(* IEC 61131-3 sources: weg-plc500-nodered-ml-pipeline/plc/src, 5 files *)

(* ---- GVL_Modbus.st ---- *)
{attribute 'qualified_only'}
VAR_GLOBAL
  (* ===================================================================== *)
  (* 1. E/S Fisicas Nativas - WEG PLC500 Local_IO (24 Vcc PNP)             *)
  (* ===================================================================== *)
  xRaw_DI0_Presenca   AT %IX0.0 : BOOL;          (* B1_SensPresenca - Contato NA *)
  xRaw_DI1_NivelAlto  AT %IX0.1 : BOOL;          (* B2_SensNivelAlto - Contato NA *)
  xRaw_DI2_Sobretemp  AT %IX0.2 : BOOL;          (* B3_SensSobretemp - Contato NA *)
  xRaw_DI3_Emergencia AT %IX0.3 : BOOL;          (* B4_Emergencia - Contato NF fail-safe (FALSE = emerg./fio partido) *)

  xDO0_Motor          AT %QX0.0 : BOOL := FALSE; (* L1_AtuMotor - LED Verde *)
  xDO1_Valvula        AT %QX0.1 : BOOL := FALSE; (* L2_AtuValvula - LED Amarelo *)
  xDO2_Alarme         AT %QX0.2 : BOOL := FALSE; (* L3_SinalAlarme - LED Vermelho *)
  xDO3_StatusOper     AT %QX0.3 : BOOL := FALSE; (* L4_StatusOper - LED Branco *)

  (* ===================================================================== *)
  (* 2. Discrete Inputs - Modbus FC02 (Enderecos base zero 0..5)           *)
  (* ===================================================================== *)
  xDI_Presenca : BOOL := FALSE; (* DI[0]: Estado filtrado (TON 50 ms) de B1_SensPresenca *)
  xDI_NivelAlto : BOOL := FALSE; (* DI[1]: Estado filtrado (TON 50 ms) de B2_SensNivelAlto *)
  xDI_Sobretemp : BOOL := FALSE; (* DI[2]: Estado filtrado (TON 50 ms) de B3_SensSobretemp *)
  xDI_EmergenciaOK : BOOL := TRUE; (* DI[3]: Estado imediato NF de B4_Emergencia (TRUE em repouso; FALSE = emergencia) *)
  xFlag_EmergTravada : BOOL := FALSE; (* DI[4]: 1 = emergencia travada aguardando rearme seguro *)
  xFlag_WatchdogAtivo : BOOL := FALSE; (* DI[5]: 1 = heartbeat estagnado > uiTimeout_WD_ms *)

  (* ===================================================================== *)
  (* 3. Coils - Modbus FC01/05/15 (Enderecos base zero 0..4)               *)
  (* ===================================================================== *)
  xCmd_Motor : BOOL := FALSE; (* Coil[0]: Comando remoto para L1_AtuMotor (DO0) *)
  xCmd_Valvula : BOOL := FALSE; (* Coil[1]: Comando remoto para L2_AtuValvula (DO1) *)
  xCmd_Alarme : BOOL := FALSE; (* Coil[2]: Comando remoto para L3_SinalAlarme (DO2) *)
  xCmd_ResetFalha : BOOL := FALSE; (* Coil[3]: Pulso de rearme (borda de subida; valido se DI3=1 e DI2=0) *)
  xCmd_HabRemoto : BOOL := FALSE; (* Coil[4]: 1 = habilita modo automatico supervisionado *)

  (* ===================================================================== *)
  (* 4. Input Registers - Modbus FC04 (Enderecos base zero 0..7)           *)
  (* ===================================================================== *)
  uiCnt_Presenca : UINT := 0; (* IR[0]: Contador modular 16 bits de B1 (0..65535) *)
  uiCnt_NivelAlto : UINT := 0; (* IR[1]: Contador modular 16 bits de B2 (0..65535) *)
  uiCnt_Sobretemp : UINT := 0; (* IR[2]: Contador modular 16 bits de B3 (0..65535) *)
  uiCnt_Emergencia : UINT := 0; (* IR[3]: Contador modular 16 bits de eventos em B4 (0..65535) *)
  uiEstado_CLP : UINT := 0; (* IR[4]: 0=INIT, 1=NORMAL_AUTO, 2=ALERTA, 3=MODO_DEGRADADO, 4=EMERGENCIA_TRAV *)
  wMascara_DO_Real : WORD := 0; (* IR[5]: Bitmask das saidas fisicas (bit0=DO0..bit3=DO3) *)
  uiEcho_Heartbeat : UINT := 0; (* IR[6]: Eco do ultimo valor de heartbeat recebido *)
  uiCod_Intertrav : UINT := 0; (* IR[7]: 0=Nenhum, 1=Emergencia, 2=Sobretemp, 3=Watchdog *)

  (* ===================================================================== *)
  (* 5. Holding Registers - Modbus FC03/06/16 (Enderecos base zero 0..3)   *)
  (* ===================================================================== *)
  uiHeartbeat_Sup : UINT := 0; (* HR[0]: Heartbeat ciclico 1..65535 (aliases de compatibilidade: uiHeartbeat_NR, uiHeartbeat_N8N) *)
  uiTimeout_WD_ms : UINT := 5000; (* HR[1]: Timeout do watchdog em ms [2000..30000], padrao 5000 *)
  uiSeveridade_IA : UINT := 0; (* HR[2]: 0=NORMAL, 1=ATENCAO, 2=CRITICO, 3=EMERGENCIA *)
  uiVersao_Mapa : UINT := 100; (* HR[3]: Versao fixa do contrato Modbus (100 = v1.0) *)
END_VAR

(* ---- FB_DebounceCounter.st ---- *)
FUNCTION_BLOCK FB_DebounceCounter
VAR_INPUT
  xRawInput       : BOOL;           (* Sinal fisico bruto (%IX0.x) *)
  xEnableDebounce : BOOL := TRUE;   (* TRUE = filtro TON (DI0..DI2); FALSE = imediato sem retardo (DI3 NF) *)
  tDebounceTime   : TIME := T#50MS; (* Tempo de estabilizacao de contato *)
  xCountOnFalling : BOOL := FALSE;  (* FALSE = borda de subida (NA); TRUE = borda de descida / NOT (NF DI3) *)
END_VAR
VAR_OUTPUT
  xFiltered       : BOOL := FALSE;  (* Estado filtrado (ou direto para DI3) *)
END_VAR
VAR_IN_OUT
  uiCounter       : UINT;           (* Contador modular 16 bits (wrap natural 65535 -> 0) *)
END_VAR
VAR
  tonDebounce     : STANDARD.TON;
  rtEdge          : STANDARD.R_TRIG;
  xEdgeSignal     : BOOL := FALSE;
END_VAR

IF xEnableDebounce THEN
  tonDebounce(IN := xRawInput, PT := tDebounceTime);
  xFiltered := tonDebounce.Q;
ELSE
  (* Entrada fail-safe DI3 atua sem retardo no primeiro ciclo de varredura *)
  xFiltered := xRawInput;
END_IF;

IF xCountOnFalling THEN
  xEdgeSignal := NOT xFiltered;
ELSE
  xEdgeSignal := xFiltered;
END_IF;

rtEdge(CLK := xEdgeSignal);
IF rtEdge.Q THEN
  uiCounter := uiCounter + 1;
END_IF;
END_FUNCTION_BLOCK

(* ---- FB_SafetyInterlock.st ---- *)
FUNCTION_BLOCK FB_SafetyInterlock
VAR_INPUT
  xDI_EmergenciaOK    : BOOL; (* DI[3]: Contato NF; FALSE = emergencia ativa / fio partido *)
  xDI_Sobretemp       : BOOL; (* DI[2]: Termostato filtrado *)
  xDI_NivelAlto       : BOOL; (* DI[1]: Nivel alto filtrado *)
  xFlag_WatchdogAtivo : BOOL; (* DI[5]: Watchdog expirado *)
  xCmd_Motor          : BOOL; (* Coil[0] *)
  xCmd_Valvula        : BOOL; (* Coil[1] *)
  xCmd_Alarme         : BOOL; (* Coil[2] *)
  xCmd_ResetFalha     : BOOL; (* Coil[3] *)
  xCmd_HabRemoto      : BOOL; (* Coil[4] *)
  uiSeveridade_IA     : UINT; (* HR[2] *)
END_VAR
VAR_OUTPUT
  xFlag_EmergTravada  : BOOL := FALSE; (* DI[4] *)
  uiEstado_CLP        : UINT := 0;     (* IR[4] *)
  uiCod_Intertrav     : UINT := 0;     (* IR[7] *)
  xDO0_Motor          : BOOL := FALSE; (* %QX0.0 *)
  xDO1_Valvula        : BOOL := FALSE; (* %QX0.1 *)
  xDO2_Alarme         : BOOL := FALSE; (* %QX0.2 *)
  xDO3_StatusOper     : BOOL := FALSE; (* %QX0.3 *)
  wMascara_DO_Real    : WORD := 0;     (* IR[5] *)
END_VAR
VAR
  rtResetFalha        : STANDARD.R_TRIG;
END_VAR

(* Deteccao de borda de subida no comando de rearme executada em todo ciclo sem mutar Coil[3] *)
rtResetFalha(CLK := xCmd_ResetFalha);

(* Travamento de emergencia fail-safe e rearme seguro *)
IF NOT xDI_EmergenciaOK THEN
  xFlag_EmergTravada := TRUE;
ELSIF xCmd_ResetFalha AND rtResetFalha.Q AND xDI_EmergenciaOK AND NOT xDI_Sobretemp THEN
  xFlag_EmergTravada := FALSE;
END_IF;

(* Maquina de estados e intertravamento local com precedencia estrita *)
IF xFlag_EmergTravada THEN
  uiEstado_CLP    := 4;
  uiCod_Intertrav := 1;
  xDO0_Motor      := FALSE;
  xDO1_Valvula    := FALSE;
  xDO2_Alarme     := TRUE;
  xDO3_StatusOper := FALSE;
ELSIF xDI_Sobretemp THEN
  uiEstado_CLP    := 2;
  uiCod_Intertrav := 2;
  xDO0_Motor      := FALSE;
  xDO1_Valvula    := TRUE;
  xDO2_Alarme     := TRUE;
  (* Reconciliacao 04_implementacao_clp.tex:141 vs :165/PROJECT.md:110: exige modo remoto ativo alem de watchdog saudavel *)
  xDO3_StatusOper := (NOT xFlag_WatchdogAtivo) AND xCmd_HabRemoto;
ELSIF xFlag_WatchdogAtivo THEN
  uiEstado_CLP    := 3;
  uiCod_Intertrav := 3;
  xDO0_Motor      := FALSE;
  xDO1_Valvula    := xDI_NivelAlto;
  xDO2_Alarme     := TRUE;
  xDO3_StatusOper := FALSE;
ELSIF xCmd_HabRemoto THEN
  uiCod_Intertrav := 0;
  uiEstado_CLP    := SEL((uiSeveridade_IA > 0) OR xDI_NivelAlto, UINT#1, UINT#2);
  xDO0_Motor      := xCmd_Motor;
  xDO1_Valvula    := xCmd_Valvula OR xDI_NivelAlto;
  xDO2_Alarme     := xCmd_Alarme OR (uiSeveridade_IA >= 2);
  xDO3_StatusOper := TRUE;
ELSE
  uiEstado_CLP    := 0;
  uiCod_Intertrav := 0;
  xDO0_Motor      := FALSE;
  xDO1_Valvula    := FALSE;
  xDO2_Alarme     := FALSE;
  xDO3_StatusOper := FALSE;
END_IF;

(* Espelhamento das saidas fisicas reais em bitmask (IR[5]) *)
wMascara_DO_Real := BOOL_TO_WORD(xDO0_Motor)
                 OR SHL(BOOL_TO_WORD(xDO1_Valvula), 1)
                 OR SHL(BOOL_TO_WORD(xDO2_Alarme), 2)
                 OR SHL(BOOL_TO_WORD(xDO3_StatusOper), 3);
END_FUNCTION_BLOCK

(* ---- FB_WatchdogHeartbeat.st ---- *)
FUNCTION_BLOCK FB_WatchdogHeartbeat
VAR_INPUT
  uiHeartbeat     : UINT;          (* HR[0]: uiHeartbeat_Sup (aliases: uiHeartbeat_NR, uiHeartbeat_N8N) *)
  uiTimeoutMs     : UINT;          (* HR[1]: uiTimeout_WD_ms [2000..30000] *)
END_VAR
VAR_OUTPUT
  uiEcho_Heartbeat    : UINT := 0;     (* IR[6]: uiEcho_Heartbeat *)
  xFlag_WatchdogAtivo : BOOL := FALSE; (* DI[5]: xFlag_WatchdogAtivo *)
  tActiveLimit        : TIME := T#5S;  (* Limiar efetivo em TIME *)
END_VAR
VAR
  tonWatchdog     : STANDARD.TON;
  uiLastHeartbeat : UINT := 0;
END_VAR

IF (uiTimeoutMs >= 2000) AND (uiTimeoutMs <= 30000) THEN
  tActiveLimit := UINT_TO_TIME(uiTimeoutMs);
ELSE
  tActiveLimit := T#5S;
END_IF;

(* Avaliar TON ANTES de atualizar uiLastHeartbeat para reiniciar por 1 ciclo na mudanca *)
tonWatchdog(
  IN := (uiHeartbeat = uiLastHeartbeat),
  PT := tActiveLimit
);

IF uiHeartbeat <> uiLastHeartbeat THEN
  uiLastHeartbeat := uiHeartbeat;
  uiEcho_Heartbeat := uiHeartbeat;
END_IF;

xFlag_WatchdogAtivo := tonWatchdog.Q;
END_FUNCTION_BLOCK

(* ---- PLC_PRG.st ---- *)
PROGRAM PLC_PRG
VAR
  fbDebPresenca : FB_DebounceCounter;
  fbDebNivel    : FB_DebounceCounter;
  fbDebTemp     : FB_DebounceCounter;
  rtEmergencia  : STANDARD.R_TRIG;
  fbWatchdog    : FB_WatchdogHeartbeat;
  fbInterlock   : FB_SafetyInterlock;
END_VAR

(* 1 & 2. Debounce (50 ms em DI0..DI2, imediato NF em DI3) e contadores modulares 16 bits *)
GVL_Modbus.xRaw_DI0_Presenca := %IX0.0;
fbDebPresenca(
  xRawInput       := %IX0.0,
  xEnableDebounce := TRUE,
  tDebounceTime   := T#50MS,
  xCountOnFalling := FALSE,
  uiCounter       := GVL_Modbus.uiCnt_Presenca
);
GVL_Modbus.xDI_Presenca := fbDebPresenca.xFiltered;

GVL_Modbus.xRaw_DI1_NivelAlto := %IX0.1;
fbDebNivel(
  xRawInput       := %IX0.1,
  xEnableDebounce := TRUE,
  tDebounceTime   := T#50MS,
  xCountOnFalling := FALSE,
  uiCounter       := GVL_Modbus.uiCnt_NivelAlto
);
GVL_Modbus.xDI_NivelAlto := fbDebNivel.xFiltered;

GVL_Modbus.xRaw_DI2_Sobretemp := %IX0.2;
fbDebTemp(
  xRawInput       := %IX0.2,
  xEnableDebounce := TRUE,
  tDebounceTime   := T#50MS,
  xCountOnFalling := FALSE,
  uiCounter       := GVL_Modbus.uiCnt_Sobretemp
);
GVL_Modbus.xDI_Sobretemp := fbDebTemp.xFiltered;

GVL_Modbus.xRaw_DI3_Emergencia := %IX0.3;
GVL_Modbus.xDI_EmergenciaOK := %IX0.3;
rtEmergencia(CLK := NOT GVL_Modbus.xDI_EmergenciaOK);
IF rtEmergencia.Q THEN
  GVL_Modbus.uiCnt_Emergencia := GVL_Modbus.uiCnt_Emergencia + 1;
END_IF;

(* 3. Supervisao de enlace Modbus TCP/IP (Watchdog via HR[0]/HR[1]) *)
fbWatchdog(
  uiHeartbeat         := GVL_Modbus.uiHeartbeat_Sup,
  uiTimeoutMs         := GVL_Modbus.uiTimeout_WD_ms,
  uiEcho_Heartbeat    => GVL_Modbus.uiEcho_Heartbeat,
  xFlag_WatchdogAtivo => GVL_Modbus.xFlag_WatchdogAtivo
);

(* 4, 5 & 6a. Travamento fail-safe, FSM com precedencia estrita e wMascara_DO_Real *)
fbInterlock(
  xDI_EmergenciaOK    := GVL_Modbus.xDI_EmergenciaOK,
  xDI_Sobretemp       := GVL_Modbus.xDI_Sobretemp,
  xDI_NivelAlto       := GVL_Modbus.xDI_NivelAlto,
  xFlag_WatchdogAtivo := GVL_Modbus.xFlag_WatchdogAtivo,
  xCmd_Motor          := GVL_Modbus.xCmd_Motor,
  xCmd_Valvula        := GVL_Modbus.xCmd_Valvula,
  xCmd_Alarme         := GVL_Modbus.xCmd_Alarme,
  xCmd_ResetFalha     := GVL_Modbus.xCmd_ResetFalha,
  xCmd_HabRemoto      := GVL_Modbus.xCmd_HabRemoto,
  uiSeveridade_IA     := GVL_Modbus.uiSeveridade_IA,
  xFlag_EmergTravada  => GVL_Modbus.xFlag_EmergTravada,
  uiEstado_CLP        => GVL_Modbus.uiEstado_CLP,
  uiCod_Intertrav     => GVL_Modbus.uiCod_Intertrav,
  xDO0_Motor          => GVL_Modbus.xDO0_Motor,
  xDO1_Valvula        => GVL_Modbus.xDO1_Valvula,
  xDO2_Alarme         => GVL_Modbus.xDO2_Alarme,
  xDO3_StatusOper     => GVL_Modbus.xDO3_StatusOper,
  wMascara_DO_Real    => GVL_Modbus.wMascara_DO_Real
);

(* Escrita direta nas saidas fisicas 24 Vcc PNP (%QX0.0..%QX0.3) *)
%QX0.0 := GVL_Modbus.xDO0_Motor;
%QX0.1 := GVL_Modbus.xDO1_Valvula;
%QX0.2 := GVL_Modbus.xDO2_Alarme;
%QX0.3 := GVL_Modbus.xDO3_StatusOper;

(* 6b. Reforco da versao do mapa Modbus a cada ciclo de 10 ms *)
GVL_Modbus.uiVersao_Mapa := 100;
END_PROGRAM
